(* IEC 61131-3 sources: plc-vscode/tests/st/all/trust-platform/crates/trust-runtime/tests/fixtures/plcopen_motion/single_axis_negative_transition_vel_zero/src, 1 file *)

(* ---- tests.st ---- *)
TEST_PROGRAM plcopen_motion_single_axis_negative_transition_vel_zero
VAR
    WrongBufferMode : MC_BUFFER_MODE;
END_VAR

WrongBufferMode := MC_BUFFER_MODE#mcTransitionVelZero;
END_TEST_PROGRAM
